{region 'Documentation'}
(*!
<summary>Compares Expected with the prefix of the selected IN range.</summary>
<description>

StartIndex is an absolute declared IN index, not an offset. Length selects 1..255
elements; the complete selected range must fit IN. Invalid references or ranges report
Error.

Keep supplied arrays stable for the call. Input data is read, not copied or retained as a
snapshot.

Comparison applies Mask to both values; bits outside it are ignored. The default mask
selects all bits.

The complete Expected pattern must be nonempty and fit the selected IN range; an
oversized pattern reports Error, not a missing-match result.

</description>
*)
{endregion}
FUNCTION_BLOCK AssertArrayStartsWithArray_Word EXTENDS AssertionBase
VAR_INPUT
    Mask : WORD := WORD#16#FFFF; //! Bits included in each element comparison.
    StartIndex : DINT; //! First index of the selected IN range.
    Length : USINT; //! Number of selected elements starting at StartIndex; must fit the array range; valid range 1..255.
END_VAR
VAR_IN_OUT CONSTANT
    IN : ARRAY[*] OF WORD; //! Read-only actual data; the selected range must remain stable during the call.
    Expected : ARRAY[*] OF WORD; //! Read-only expected sequence starting at its own lower bound; must fit the selected actual range.
END_VAR

SUPER^();

{region 'Documentation'}
(*!
<summary>Validate the selected range and expectations before comparing elements.</summary>
*)
{endregion}
METHOD PROTECTED Assert
VAR
    InLowerIndex : DINT;
    InUpperIndex : DINT;
    ExpectedLowerIndex : DINT;
    ExpectedUpperIndex : DINT;
    ExpectedLength : LINT;
    EndIndex : LINT;
    Offset : LINT;
    InIndex : DINT;
    ExpectedIndex : DINT;
    Message : STRING(GVL_Constants.MessageLength);
    ExpectedText : STRING(GVL_Constants.AssertionValueLength);
    ActualText : STRING(GVL_Constants.AssertionValueLength);
END_VAR
VAR CONSTANT
    HexDigitCount : USINT := 4;
END_VAR
IF NOT EvaluationActive THEN
    RETURN;
END_IF;

IF Result = E_Result.Error THEN
    RETURN;
END_IF;

// C0371: FB inputs are checked here before any reference access.
{warning disable C0371}
IF NOT __ISVALIDREF(IN) THEN
    Error(Message := 'Assertion error: IN reference is invalid.');
    RETURN;
END_IF;

IF NOT __ISVALIDREF(Expected) THEN
    Error(Message := 'Assertion error: Expected reference is invalid.');
    RETURN;
END_IF;

InLowerIndex := LOWER_BOUND(IN, 1);
InUpperIndex := UPPER_BOUND(IN, 1);
ExpectedLowerIndex := LOWER_BOUND(Expected, 1);
ExpectedUpperIndex := UPPER_BOUND(Expected, 1);
ExpectedLength := DINT_TO_LINT(ExpectedUpperIndex) - DINT_TO_LINT(ExpectedLowerIndex) + 1;
EndIndex := DINT_TO_LINT(StartIndex) + USINT_TO_LINT(Length) - 1;

IF (Length = 0) OR (ExpectedLength <= 0)
    OR (ExpectedLength > USINT_TO_LINT(Length))
    OR (StartIndex < InLowerIndex) OR (StartIndex > InUpperIndex)
    OR (EndIndex > DINT_TO_LINT(InUpperIndex)) THEN
    Message := CONCAT('Assertion error: array range is invalid. StartIndex = ',
        DINT_TO_STRING(StartIndex));
    Message := CONCAT(Message, ', EndIndex = ');
    Message := CONCAT(Message, LINT_TO_STRING(EndIndex));
    Message := CONCAT(Message, ', InLowerIndex = ');
    Message := CONCAT(Message, DINT_TO_STRING(InLowerIndex));
    Message := CONCAT(Message, ', InUpperIndex = ');
    Message := CONCAT(Message, DINT_TO_STRING(InUpperIndex));
    Message := CONCAT(Message, ', ExpectedLength = ');
    Message := CONCAT(Message, LINT_TO_STRING(ExpectedLength));
    Message := CONCAT(Message, '.');
    Error(Message := Message);
    RETURN;
END_IF;

IF Result = E_Result.Failed THEN
    RETURN;
END_IF;

FOR Offset := 0 TO ExpectedLength - 1 DO
    InIndex := LINT_TO_DINT(DINT_TO_LINT(StartIndex) + Offset);
    ExpectedIndex := LINT_TO_DINT(DINT_TO_LINT(ExpectedLowerIndex) + Offset);
    IF (IN[InIndex] AND Mask) <> (Expected[ExpectedIndex] AND Mask) THEN
        ExpectedText := CreateAssertionTextValue_Hex(Value := WORD_TO_LWORD(Expected[ExpectedIndex]),
            DigitCount := HexDigitCount);
        ActualText := CreateAssertionTextValue_Hex(Value := WORD_TO_LWORD(IN[InIndex]),
            DigitCount := HexDigitCount);
        Message := CONCAT('Assertion failed: array prefix differs. Expected[',
            DINT_TO_STRING(ExpectedIndex));
        Message := CONCAT(Message, '] = ');
        Message := CONCAT(Message, ExpectedText);
        Message := CONCAT(Message, ', IN[');
        Message := CONCAT(Message, DINT_TO_STRING(InIndex));
        Message := CONCAT(Message, '] = ');
        Message := CONCAT(Message, ActualText);
        Message := CONCAT(Message, '.');
        Message := CONCAT(Message, ' Mask = ');
        Message := CONCAT(Message, CreateAssertionTextValue_Hex(Value := WORD_TO_LWORD(Mask),
            DigitCount := HexDigitCount));
        Fail(Message := Message);
        RETURN;
    END_IF;
END_FOR;

Pass();
{warning restore C0371}
END_METHOD

END_FUNCTION_BLOCK

(* stored: Version 1.1.0.1
   POU AssertArrayStartsWithArray_Word: Id {87c7e592-4033-4021-bb12-da2b20227f8e}, SpecialFunc None
   Folder Internal: Id {59b26f99-ba8b-4be5-a4d5-ec6d02b337b8}
   Method Assert: Id {55d3386b-9155-4a2f-875c-1924fd492b11} *)
